(*
SPDX-FileCopyrightText: © 2026 Oleksandr Tiutyk <trofimich@gmail.com>
SPDX-License-Identifier: MIT
License: https://opensource.org/license/mit
*)

(*!
<summary>Groups the seven independent queue cleanup cases.</summary>
<description>
Owns the cases and their fixed child array for single-task use. Copying invalidates the child bindings.
</description>
*)

{attribute 'no_assign'}
{attribute 'no_explicit_call' := 'do not call this function block directly'}
FUNCTION_BLOCK TaskQueueCleanupTestGroup EXTENDS TOF_Testing.TestGroup<7>
VAR_STAT
	{attribute 'hide'}
	_ClassName : STRING := __POUNAME();
END_VAR
VAR
	_DelayedCleanupAndReuse : TaskQueueCleanupScenarioTest(
		name := "DelayedCleanupAndReuse",
		parent := THIS^,
		scenario := QUEUE_CLEANUP_TEST_SCENARIO.DELAYED_CLEANUP_AND_REUSE
	);
	_RepeatedExecuteFailure : TaskQueueCleanupScenarioTest(
		name := "RepeatedExecuteFailure",
		parent := THIS^,
		scenario := QUEUE_CLEANUP_TEST_SCENARIO.REPEATED_EXECUTE_FAILURE
	);
	_CancelRequestFailure : TaskQueueCleanupScenarioTest(
		name := "CancelRequestFailure",
		parent := THIS^,
		scenario := QUEUE_CLEANUP_TEST_SCENARIO.CANCEL_REQUEST_FAILURE
	);
	_MessageFormattingFailure : TaskQueueCleanupScenarioTest(
		name := "MessageFormattingFailure",
		parent := THIS^,
		scenario := QUEUE_CLEANUP_TEST_SCENARIO.MESSAGE_FORMATTING_FAILURE
	);
	_ExternalCancelDuringCleanup : TaskQueueCleanupScenarioTest(
		name := "ExternalCancelDuringCleanup",
		parent := THIS^,
		scenario := QUEUE_CLEANUP_TEST_SCENARIO.EXTERNAL_CANCEL_DURING_CLEANUP
	);
	_HeldCleanup : TaskQueueCleanupScenarioTest(
		name := "HeldCleanup",
		parent := THIS^,
		scenario := QUEUE_CLEANUP_TEST_SCENARIO.HELD_CLEANUP
	);
	_ExternalCancelWithReleaseFailure : TaskQueueCleanupScenarioTest(
		name := "ExternalCancelWithReleaseFailure",
		parent := THIS^,
		scenario := QUEUE_CLEANUP_TEST_SCENARIO.EXTERNAL_CANCEL_WITH_RELEASE_FAILURE
	);

	_Children : ARRAY [0.._ChildCount - 1] OF TOF_Testing.ITestElement :=
	[
		_DelayedCleanupAndReuse,
		_RepeatedExecuteFailure,
		_CancelRequestFailure,
		_MessageFormattingFailure,
		_ExternalCancelDuringCleanup,
		_HeldCleanup,
		_ExternalCancelWithReleaseFailure
	];
END_VAR

//! <summary>Borrows the fixed child array. Callers must not modify it.</summary>
{attribute 'monitoring' := 'call'}
PROPERTY Children : REFERENCE TO ARRAY [0.._ChildCount - 1] OF TOF_Testing.ITestElement
GET
Children REF= _Children;
END_GET
END_PROPERTY

//! <summary>Borrows the concrete class name. Callers must not modify it.</summary>
{attribute 'monitoring' := 'call'}
PROPERTY ClassName : REFERENCE TO STRING
GET
ClassName REF= _ClassName;
END_GET
END_PROPERTY

//! <summary>Borrows the compiler-initialized namespace name. Callers must not modify it.</summary>
{attribute 'monitoring' := 'call'}
PROPERTY NamespaceName : REFERENCE TO STRING
GET
NamespaceName REF= CurrentNamespace.Name;
END_GET
END_PROPERTY

//! <summary>Reports the complete concrete instance size in bytes.</summary>
{attribute 'monitoring' := 'call'}
PROPERTY SelfSize : ULINT
GET
SelfSize := XSIZEOF(THIS^);
END_GET
END_PROPERTY

END_FUNCTION_BLOCK

(* stored: Version 1.1.0.1
   POU TaskQueueCleanupTestGroup: Id {6c703de6-c8b2-4802-a488-37740853b79f}, SpecialFunc None
   Property Children: Id {585f2d0c-1105-49d5-bc3e-79adc2b63f9c}
   Get Get: Id {d50f7e2d-0e3f-48fe-92ab-1daa27fc95a1}
   Property ClassName: Id {35e88aa5-dff8-43c4-81dc-2ffd699c9fca}
   Get Get: Id {dd2f954a-2daf-4066-8d3d-07add2d734ee}
   Property NamespaceName: Id {ac9dc1d4-9bd1-476d-9c94-c1924468ded4}
   Get Get: Id {614c477c-afa3-4a90-ad33-f6b4ecf8086b}
   Property SelfSize: Id {cdfedb02-6947-412c-9aa1-a8ee5671d2c2}
   Get Get: Id {608b0fe3-6a8c-49d4-a073-76c0feecdca2} *)
